{region 'Documentation'}
(*!
<summary>Assertion-specific identity and result view; initialization remains an instance API.</summary>
*)
{endregion}
INTERFACE I_Assertion EXTENDS I_ResultProvider

END_INTERFACE

(* stored: Version 1.1.0.1
   Itf I_Assertion: Id {69c8dce9-9b31-45d4-b6d1-94dd1e4c8ab9} *)
